(* IEC 61131-3 sources: llm-plc-st-eval/data/definitivo/gemini-3.1-pro-preview/I1/few_shot, 3 files *)

(* ---- ejec_1.st ---- *)
FUNCTION_BLOCK FB_Semaforo
VAR_INPUT
    habilitado : BOOL; (* Habilitacion del semaforo *)
END_VAR
VAR_OUTPUT
    luzV : BOOL; (* Luz verde *)
    luzA : BOOL; (* Luz amarilla *)
    luzR : BOOL; (* Luz roja *)
END_VAR
VAR
    estado : INT := 0; (* 0: Verde, 1: Amarillo, 2: Rojo *)
    tFase : TON; (* Temporizador para las fases del semaforo *)
    tParpadeo : TON; (* Temporizador para el parpadeo *)
    estadoBlink : BOOL := TRUE; (* Estado de la luz intermitente *)
END_VAR

IF habilitado THEN
    (* Secuencia normal del semaforo *)
    CASE estado OF
        0: tFase(IN := TRUE, PT := T#20S); (* Verde *)
        1: tFase(IN := TRUE, PT := T#4S);  (* Amarillo *)
        2: tFase(IN := TRUE, PT := T#15S); (* Rojo *)
    END_CASE;

    (* Cambio de fase al terminar el tiempo *)
    IF tFase.Q THEN
        estado := (estado + 1) MOD 3;
        tFase(IN := FALSE); (* Reiniciar temporizador para la siguiente fase *)
    END_IF;

    (* Asignacion de salidas *)
    luzV := (estado = 0);
    luzA := (estado = 1);
    luzR := (estado = 2);

    (* Reiniciar variables del modo intermitente *)
    tParpadeo(IN := FALSE);
    estadoBlink := TRUE;
ELSE
    (* Modo deshabilitado: Amarillo intermitente *)
    estado := 0; (* Preparar reinicio en verde *)
    tFase(IN := FALSE); (* Reiniciar temporizador de secuencia *)

    (* Generador de pulsos de 1 segundo *)
    tParpadeo(IN := TRUE, PT := T#1S);
    IF tParpadeo.Q THEN
        estadoBlink := NOT estadoBlink;
        tParpadeo(IN := FALSE); (* Reiniciar temporizador de parpadeo *)
    END_IF;

    (* Asignacion de salidas *)
    luzV := FALSE;
    luzR := FALSE;
    luzA := estadoBlink;
END_IF;
END_FUNCTION_BLOCK

(* ---- ejec_2.st ---- *)
FUNCTION_BLOCK FB_Semaforo
VAR_INPUT
    habilitado : BOOL; (* Habilitacion del semaforo *)
END_VAR
VAR_OUTPUT
    luzV : BOOL; (* Luz verde *)
    luzA : BOOL; (* Luz amarilla *)
    luzR : BOOL; (* Luz roja *)
END_VAR
VAR
    estado : INT := 0; (* 0: Intermitente, 1: Verde, 2: Amarillo, 3: Rojo *)
    tSecuencia : TON;  (* Temporizador para la secuencia normal *)
    tBlink1 : TON;     (* Temporizador 1 para parpadeo (tiempo encendido) *)
    tBlink2 : TON;     (* Temporizador 2 para parpadeo (tiempo apagado) *)
    tiempoActual : TIME;
    transicion : BOOL;
END_VAR

(* Control de estado principal *)
IF NOT habilitado THEN
    estado := 0;
ELSIF estado = 0 THEN
    estado := 1; (* Reinicia en verde al habilitarse *)
END_IF;

(* Asignacion de tiempos y luces segun el estado *)
CASE estado OF
    0: (* Amarillo intermitente *)
        luzV := FALSE;
        luzA := NOT tBlink1.Q;
        luzR := FALSE;
    1: (* Verde *)
        tiempoActual := T#20S;
        luzV := TRUE;
        luzA := FALSE;
        luzR := FALSE;
    2: (* Amarillo *)
        tiempoActual := T#4S;
        luzV := FALSE;
        luzA := TRUE;
        luzR := FALSE;
    3: (* Rojo *)
        tiempoActual := T#15S;
        luzV := FALSE;
        luzA := FALSE;
        luzR := TRUE;
END_CASE;

(* Actualizacion de temporizadores *)
tSecuencia(IN := habilitado AND NOT transicion, PT := tiempoActual);
transicion := tSecuencia.Q;

tBlink1(IN := (estado = 0) AND NOT tBlink2.Q, PT := T#1S);
tBlink2(IN := tBlink1.Q, PT := T#1S);

(* Transiciones de la secuencia normal *)
IF transicion THEN
    CASE estado OF
        1: estado := 2;
        2: estado := 3;
        3: estado := 1;
    END_CASE;
END_IF;
END_FUNCTION_BLOCK

(* ---- ejec_3.st ---- *)
```iecst
FUNCTION_BLOCK FB_Semaforo
VAR_INPUT
    habilitado : BOOL; (* Habilita la secuencia normal *)
END_VAR
VAR_OUTPUT
    luzV : BOOL; (* Luz verde *)
    luzA : BOOL; (* Luz amarilla *)
    luzR : BOOL; (* Luz roja *)
END_VAR
VAR
    estado : INT := 0; (* 0: Verde, 1: Amarillo, 2: Rojo *)
    tVerde : TON;      (* Temporizador luz verde *)
    tAmarillo : TON;   (* Temporizador luz amarilla *)
    tRojo : TON;       (* Temporizador luz roja *)
    tBlink1 : TON;     (* Temporizador intermitencia ON *)
    tBlink2 : TON;     (* Temporizador intermitencia OFF *)
END_VAR

(* Control de estados y reinicio *)
IF NOT habilitado THEN
    estado := 0; (* Reinicia la secuencia a verde si se deshabilita *)
ELSIF estado = 0 AND tVerde.Q THEN
    estado := 1;
ELSIF estado = 1 AND tAmarillo.Q THEN
    estado := 2;
ELSIF estado = 2 AND tRojo.Q THEN
    estado := 0;
END_IF;

(* Temporizadores de la secuencia normal *)
tVerde(IN := habilitado AND (estado = 0), PT := T#20S);
tAmarillo(IN := habilitado AND (estado = 1), PT := T#4S);
tRojo(IN := habilitado AND (estado = 2), PT := T#15S);

(* Temporizadores del modo intermitente (1s ON / 1s OFF) *)
tBlink1(IN := NOT habilitado AND NOT tBlink2.Q, PT := T#1S);
tBlink2(IN := tBlink1.Q, PT := T#1S);

(* Asignacion de salidas *)
luzV := habilitado AND (estado = 0);
luzR := habilitado AND (estado = 2);
luzA := (habilitado AND (estado = 1)) OR (NOT habilitado AND NOT tBlink1.Q);

END_FUNCTION_BLOCK
```
